(* IEC 61131-3 sources: SRCI_CLIENT_PLC/RobotLibrary/Library/POUs/Write/MC_WriteRobotReferenceDynamics/Structures, 4 files *)

(* ---- WriteRobotReferenceDynamicsOutCmd.st ---- *)
{attribute 'pack_mode' := '1'}
// -------------------------------------------------------------------------
//  SRCI Robot Library
// -------------------------------------------------------------------------
//
//  Object:      WriteRobotReferenceDynamicsOutCmd
//  Author:      Thorsten Brach
//  Date:        2024-08-08
//
//  Description:
//
//
//  Copyright:
//    (C) 2024 Thorsten Brach. All rights reserved
//             Licensed under the MIT License.
//
//  Disclaimer:
//    This project is provided without any guarantee and can be used for
//    private and commercial purposes. Any use is at the user’s
//    own risk and responsibility.
//
// -------------------------------------------------------------------------
TYPE WriteRobotReferenceDynamicsOutCmd :
STRUCT
  /// Commanded reference dynamics values according to Table 6-158
  ReferenceDynamicValues : ReferenceDynamics;
END_STRUCT
END_TYPE

(* ---- WriteRobotReferenceDynamicsParCmd.st ---- *)
{attribute 'pack_mode' := '1'}
// -------------------------------------------------------------------------
//  SRCI Robot Library
// -------------------------------------------------------------------------
//
//  Object:      WriteRobotReferenceDynamicsParCmd
//  Author:      Thorsten Brach
//  Date:        2024-08-08
//
//  Description:
//
//
//  Copyright:
//    (C) 2024 Thorsten Brach. All rights reserved
//             Licensed under the MIT License.
//
//  Disclaimer:
//    This project is provided without any guarantee and can be used for
//    private and commercial purposes. Any use is at the user’s
//    own risk and responsibility.
//
// -------------------------------------------------------------------------
TYPE WriteRobotReferenceDynamicsParCmd :
STRUCT
  /// Reference dynamics values according TO Table 6-158.
  DynamicValues : ReferenceDynamics := ( VelocityReference := -1.0, AccelerationReference := -1.0, DecelerationReference := -1.0, JerkReference := -1.0); // ST-FIX F126: spec 6.2.13 / 6.2.14: input of the write command, default '<0' = do not change; 0.0 wrote 0 (minimum) for every value that was not set
END_STRUCT
END_TYPE

(* ---- WriteRobotReferenceDynamicsRecvData.st ---- *)
{attribute 'pack_mode' := '1'}
// -------------------------------------------------------------------------
//  SRCI Robot Library
// -------------------------------------------------------------------------
//
//  Object:      WriteRobotReferenceDynamicsRecvData
//  Author:      Thorsten Brach
//  Date:        2024-08-08
//
//  Description:
//
//
//  Copyright:
//    (C) 2024 Thorsten Brach. All rights reserved
//             Licensed under the MIT License.
//
//  Disclaimer:
//    This project is provided without any guarantee and can be used for
//    private and commercial purposes. Any use is at the user’s
//    own risk and responsibility.
//
// -------------------------------------------------------------------------
TYPE WriteRobotReferenceDynamicsRecvData EXTENDS RspHeader :
STRUCT
  /// Commanded reference dynamics values according to Table 6-158
  ReferenceDynamicValues : ReferenceDynamics;
END_STRUCT
END_TYPE

(* ---- WriteRobotReferenceDynamicsSendData.st ---- *)
{attribute 'pack_mode' := '1'}
// -------------------------------------------------------------------------
//  SRCI Robot Library
// -------------------------------------------------------------------------
//
//  Object:      WriteRobotReferenceDynamicsSendData
//  Author:      Thorsten Brach
//  Date:        2024-08-08
//
//  Description:
//
//
//  Copyright:
//    (C) 2024 Thorsten Brach. All rights reserved
//             Licensed under the MIT License.
//
//  Disclaimer:
//    This project is provided without any guarantee and can be used for
//    private and commercial purposes. Any use is at the user’s
//    own risk and responsibility.
//
// -------------------------------------------------------------------------
TYPE WriteRobotReferenceDynamicsSendData EXTENDS CmdHeader:
STRUCT

  DynamicValues : ReferenceDynamics;
(*
  /// Timestamp
  Timestamp             : IEC_TIMESTAMP;
  /// Path velocity [mm/s](tangent) at 100%
  /// • <0: (default) - Do not change values
  /// • ≥0: Change values according to input value
  VelocityReference     : UINT;
  /// Path acceleration [mm/s2] at 100%
  /// • <0: (default) - Do not change values
  /// • ≥0: Change values according to input value
  AccelerationReference : UINT;
  /// Path deceleration [mm/s2] at 100%
  /// • <0: (default) - Do not change values
  /// • ≥0: Change values according to input value
  DecelerationReference : UINT;
  /// Jerk [mm/s3] at 100%
  /// • <0: (default) - Do not change values
  /// • ≥0: Change values according to input value
  JerkReference        : UINT;
*)
END_STRUCT
END_TYPE
